// TIA Portal V21 export
// export: Created 2026-10-12T12:46:19.0678456Z, ExportSetting WithDefaults, DisplayName Totally Integrated Automation Portal, DisplayVersion V21, DisplayName STEP 7 Professional, DisplayVersion V21, DisplayName STEP 7 Safety, DisplayVersion V21, DisplayName Tech WebApplication, DisplayVersion V21, DisplayName WinCC Basic/Comfort/Advanced, DisplayVersion V21, DisplayName WinCC Unified, DisplayVersion V21
TextList "MODE"  ListRange=Bit
  TextListEntry   EntryType=SingleValue, Text="MANUAL"
  TextListEntry   EntryType=SingleValue, From=1, To=1, Text="AUTO"
